TYPE "DT_REGULATOR_VALUES_INTERFACE"
VERSION : 0.1
   STRUCT
      SCALED_REFERENCE : Real;   // SCALED REFERENCE
      OUT : Real;   // REGULATOR_OUTPUT
      SCALED_MEAS : Real;   // MEASUREMENT
   END_STRUCT;

END_TYPE

